(* IEC 61131-3 sources: axsharp/src/ix.blazor/tests/sandbox/ax-blazor-example/src, 40 files *)

(* ---- enumStationStatus.st ---- *)
TYPE enumStationStatus :
    (
        Unknown,
        Available,
        UnAvailable
    );
    END_TYPE

(* ---- stTestEnum.st ---- *)
TYPE stTestEnum :
    (
        Unknown,
        Available,
        UnAvailable
    );
END_TYPE

(* ---- CU00x.st ---- *)
CLASS CU00x EXTENDS CUBase
    VAR PUBLIC
        _cuName: STRING;
    END_VAR
END_CLASS

CLASS CUBase
    VAR PUBLIC
        _baseName : STRING;
    END_VAR
END_CLASS

(* ---- fbWorldWeatherWatch.st ---- *)
CLASS fbWorldWeatherWatch
    VAR PUBLIC
        {#ix-attr:[Container(Layout.Stack)]}
        {#ix-set:AttributeName = "North pole station"}
        //{#ix-set:OpenMap = "https://www.openstreetmap.org/?mlat=74.652&mlon=-95.556#map=6/74.652/-95.556"}
        NorthPole : structWeatherStation := (StationICAO := 'CYRB');
        {#ix-attr:[Container(Layout.Stack)]}
        {#ix-set:AttributeName = "South pole station"}
        //{#ix-set:OpenMap = "https://www.openstreetmap.org/?mlat=-85.05113&mlon=-16.80701#map=1/-85.05113/-16.80701"}
        SouthPole : structWeatherStation := (StationICAO := 'NZSP');
        {#ix-attr:[Container(Layout.Stack)]}
        {#ix-set:AttributeName = "Verl, Germany"}
        //{#ix-set:OpenMap = "https://www.openstreetmap.org/?mlat=51.5799&mlon=8.415#map=6/51.5799/8.4155"}
        Verl : structWeatherStation := (StationICAO := 'EDLP');
        {#ix-attr:[Container(Layout.Stack)]}
        {#ix-set:AttributeName = "Kriva, Slovakia"}
        //{#ix-set:OpenMap = "https://www.openstreetmap.org/?mlat=48.1723&mlon=17.2158#map=6/48.1723/17.2158"}
        Kriva : structWeatherStation := (StationICAO := 'LZIB');
    END_VAR

END_CLASS

(* ---- GroupBox_other.st ---- *)
CLASS GroupBox_other
    VAR PUBLIC
        {#ix-set:AttributeName = "B1"}
        B1: INT;

        {#ix-attr:[Container(Layout.Stack)]}
        {#ix-set:AttributeName = "B2"}
        B2: INT;

        {#ix-attr:[Container(Layout.Stack)]}
        {#ix-set:AttributeName = "A1"}
        Piston_A1 : STRING;
        {#ix-set:AttributeName = "A2"}
        Piston_A2 : STRING;
        {#ix-set:AttributeName = "A3"}
        Piston_A3 : STRING;
        {#ix-set:AttributeName = "A4"}
        Piston_A4 : STRING;

        {#ix-attr:[Container(Layout.Tabs)]}
        Piston_A21 : INT;
        {#ix-set:AttributeName = "A5"}
        Piston_A22 : INT;
        {#ix-set:AttributeName = "A6"}
        Piston_A23 : INT;
        {#ix-set:AttributeName = "A7"}
        Piston_A24 : INT;

        {#ix-attr:[Container(Layout.UniformGrid)]}
        Piston_A31 : REAL;
        {#ix-set:AttributeName = "A8"}
        Piston_A32 : REAL;
        {#ix-set:AttributeName = "A9"}
        Piston_A33 : REAL;
        {#ix-set:AttributeName = "A10"}
        Piston_A34 : REAL;

        Piston_A41 : BOOL;
        {#ix-set:AttributeName = "A11"}
        Piston_A42 : BOOL;
        {#ix-set:AttributeName = "A12"}
        Piston_A43 : BOOL;
        {#ix-set:AttributeName = "A13"}
        Piston_A44 : BOOL;
        {#ix-set:AttributeName = "Servo S1"}
        Servo_S1: TestStructOneGroupWithLayout;
        {#ix-attr:[Container(Layout.Stack)]}
        {#ix-set:AttributeName = "ABB S2"}
        Servo_S2: STRING;
    END_VAR

END_CLASS

(* ---- MAIN.st ---- *)
CLASS MAIN
    VAR PUBLIC
        {#ix-set:AttributeName = "<#Hello#> <#World#>"}
        Hello_World : STRING := 'Hello world!';
        {#ix-set:AttributeName = "cislo"}
        cislo : INT;
        {#ix-set:AttributeName = "bool_val"}
        boolValue : BOOL;
        {#ix-set:AttributeName = "Position"}
        Position : LREAL;
        {#ix-set:AttributeName = "Struct"}
        instanceOfstTest: stTest;
        {#ix-set:AttributeName = "Struct2"}
        instanceOfstTest2: stTest2 ;
        {#ix-set:AttributeName = "instanceOfStTest3"}
        instanceOfstTest3: stTest3 ;
        {#ix-set:AttributeName = "BlazorStruct"}
        instanceOfstBlazor: stBlazor := (testInteger := 10, testString := 'ahoj');
        arr1 : ARRAY [0..2] OF stTest := [(p1 := 6, p2 := 3),(p1 := 9, p2 := 10),(p1 := 12,p2 := 33)];
        arr2 :ARRAY [0..5] OF INT;
        dateVar : DATE;

        {#ix-set:AttributeName = "instanceOfComplex"}
        instanceOfstComplex: stComplex ;
        {#ix-set:AttributeName = "instanceOfStPrimitive"}
        instanceOfstPrimitive: stTestPrimitive ;

    //	{#ix [Container(Layout.Stack)]}
        instanceOfstMultipleLayouts: stMultipleLayouts ;
        instanceOfstMultipleLayouts2: stLayouts ;

        {#ix-set:AttributeName = "instanceOfIxComponent"}
        instanceOfIxComponent: IxComponent ;

        groupBox_test: GroupBox_other;
        cu00: CU00x;
        cuBase: CUBase;
    END_VAR

END_CLASS

(* ---- prgWeatherStations.st ---- *)
{#ix-attr:[Container(Layout.Stack)]}
CLASS prgWeatherStations
    VAR PUBLIC
        {#ix-attr:[Container(Layout.Tabs)]}
        {#ix-set:AttributeName = "Weather Cyclic"}
        _weatherStations : fbWorldWeatherWatch;
        {#ix-attr:[Container(Layout.Stack)]}
        {#ix-attr:[Group(GroupLayout.GroupBox)]}
        {#ix-set:AttributeName = "What plc says"}
        PlcCommentOnCurrentWeather : STRING[254] := 'TEST';
    END_VAR
END_CLASS

(* ---- stBlazor.st ---- *)
CLASS stBlazor
    VAR PUBLIC
        {#ix-set:AttributeName = "<#Integer From PLC#>"}
        testInteger : INT;
        {#ix-set:AttributeName = "testEnum"}
        testEnum : stTestEnum;
        {#ix-set:AttributeName = "<#String From PLC#>"}
        testString : STRING;
        testReal : REAL := REAL#592.25;
        {#ix-attr:[RenderIgnore("Display")]}
        testLReal : LREAL := 42.2;
        testBool : BOOL;
        {#ix-set:AttributeName = "Complex"}
        {#ix-attr:[RenderIgnore()]}
        complexInstance : stComplex := (stComplexInteger := 33, stComplexString := 'hello world');
        {#ix-set:AttributeName = "testInstance1"}
        testInstance : stTest3;
        {#ix-set:AttributeName = "testInstance2"}
        testInstance2 : stTest3;
        {#ix-set:AttributeName = "testInstance3"}
        testInstance3 : stTest;
    END_VAR

END_CLASS

(* ---- stComplex.st ---- *)
CLASS stComplex
    VAR PUBLIC
        {#ix-set:AttributeName = "<#Integer From PLC#>"}
        stComplexInteger : INT;
        {#ix-set:AttributeName = "<#String From PLC#>"}
        stComplexString : STRING;
    END_VAR

END_CLASS

(* ---- stComplexUnknown.st ---- *)
CLASS stComplexUnknown
    VAR PUBLIC
        {#ix-set:AttributeName = "<#String unknown From PLC#>"}
        stComplexUnknownString : STRING;
        {#ix-set:AttributeName = "<#BOOL unknown From PLC#>"}
        testBool : BOOL;
        {#ix-set:AttributeName = "<#Integer unknown From PLC#>"}
        stComplexUnknowInteger : INT;
        {#ix-set:AttributeName = "<#DATE unknown From PLC#>"}
        TestDate : DATE;
    END_VAR
END_CLASS

(* ---- stExample.st ---- *)
CLASS stExample
    VAR PUBLIC
        {#ix-attr:[Container(Layout.Tabs)]}
        {#ix-attr:[Group(GroupLayout.GroupBox)]}
        {#ix-set:AttributeName = "Group name"}
        testInteger : INT;
        testEnum : stTestEnum;
        testString : STRING := 'Hello World';
        testBool : BOOL;
    END_VAR

END_CLASS

(* ---- stLayouts.st ---- *)
CLASS stLayouts
    VAR
        {#ix-set:AttributeName = "B1"}
	B1: INT;

	{#ix-attr:[Container(Layout.Stack)]}
	{#ix-set:AttributeName = "B2"}
	B2: INT;

	{#ix-attr:[Container(Layout.Stack)]}
	{#ix-set:AttributeName = "A1"}
	Piston_A1 : STRING;
	{#ix-set:AttributeName = "A2"}
	Piston_A2 : STRING;
	{#ix-set:AttributeName = "A3"}
	Piston_A3 : STRING;
	{#ix-set:AttributeName = "A4"}
	Piston_A4 : STRING;

	{#ix-attr:[Container(Layout.Tabs)]}
	Piston_A21 : INT;
	{#ix-set:AttributeName = "A5"}
	Piston_A22 : INT;
	{#ix-set:AttributeName = "A6"}
	Piston_A23 : INT;
	{#ix-set:AttributeName = "A7"}
	Piston_A24 : INT;

	{#ix-attr:[Container(Layout.UniformGrid)]}
	Piston_A31 : REAL;
	{#ix-set:AttributeName = "A8"}
	Piston_A32 : REAL;
	{#ix-set:AttributeName = "A9"}
	Piston_A33 : REAL;
	{#ix-set:AttributeName = "A10"}
	Piston_A34 : REAL;

	Piston_A41 : BOOL;
	{#ix-set:AttributeName = "A11"}
	Piston_A42 : BOOL;
	{#ix-set:AttributeName = "A12"}
	Piston_A43 : BOOL;
	{#ix-set:AttributeName = "A13"}
	Piston_A44 : BOOL;

	{#ix-set:AttributeName = "Servo S1"}
	Servo_S1: TestStructOneGroupWithLayout;
	{#ix-attr:[Container(Layout.Stack)]}
	{#ix-set:AttributeName = "ABB S2"}
	Servo_S2: STRING;
    END_VAR
END_CLASS

(* ---- stMultipleLayouts.st ---- *)
CLASS stMultipleLayouts
    VAR PUBLIC
        {#ix-attr:[Container(Layout.Tabs)]}
        {#ix-set:AttributeName = "With One Group Layout"}
        Servo_S5: TestStructOneGroupWithLayout;

        {#ix-attr:[Container(Layout.Tabs)]}
        {#ix-set:AttributeName = "Without Group Layout"}
        Servo_S6: TestStruct;

        {#ix-attr:[Container(Layout.Tabs)]}
        {#ix-set:AttributeName = "With Multiple Groups "}
        Servo_S7: TestStructMultipleGroups;

        {#ix-attr:[Container(Layout.Tabs)]}
        {#ix-set:AttributeName = "TestStruct With Main Layout  "}
        Servo_S8: TestStructWithMainLayout;

        {#ix-attr:[Container(Layout.Stack)]}
        {#ix-set:AttributeName = "A1"}
        Piston_A1 : STRING;
        {#ix-set:AttributeName = "A2"}
        Piston_A2 : STRING;
        {#ix-set:AttributeName = "A3"}
        Piston_A3 : STRING;
        {#ix-set:AttributeName = "A4"}
        Piston_A4 : STRING;

        {#ix-attr:[Container(Layout.Wrap)]}
        {#ix-set:AttributeName = "A5"}
        Piston_A21 : INT;
        {#ix-set:AttributeName = "A6"}
        Piston_A22 : INT;
        {#ix-set:AttributeName = "A7"}
        Piston_A23 : INT;
        {#ix-set:AttributeName = "A8"}
        Piston_A24 : INT;

        {#ix-attr:[Container(Layout.Tabs)]}
        Piston_A31 : REAL;
        {#ix-set:AttributeName = "A8"}
        Piston_A32 : REAL;
        {#ix-set:AttributeName = "A9"}
        Piston_A33 : REAL;
        {#ix-set:AttributeName = "A10"}
        Piston_A34 : REAL;

        {#ix-attr:[Container(Layout.UniformGrid)]}
        Piston_A41 : BOOL;
        {#ix-set:AttributeName = "A11"}
        Piston_A42 : BOOL;
        {#ix-set:AttributeName = "A12"}
        Piston_A43 : BOOL;
        {#ix-set:AttributeName = "A13"}
        Piston_A44 : BOOL;

        {#ix-attr:[Container(Layout.Stack)]}
        {#ix-set:AttributeName = "Servo S1"}
        Servo_S1: STRING;

        {#ix-attr:[Container(Layout.Stack)]}
        {#ix-set:AttributeName = "ABB S2"}
        Servo_S2: STRING;

        {#ix-attr:[Container(Layout.Tabs)]}
        {#ix-set:AttributeName = "My ix component"}
        component: IxComponent;
        {#ix-set:AttributeName = "Servo S3"}
        Servo_S3: stTest3;
        {#ix-set:AttributeName = "Servo S4"}
        Servo_S4: stTest3;

    END_VAR

END_CLASS

(* ---- structWeatherStation.st ---- *)
CLASS structWeatherStation
    VAR PUBLIC
        {#ix-set:AttributeName = "Station name (ICAO)"}
        StationICAO : STRING[4];
        {#ix-set:AttributeName = "Station status"}
        StationStatus : enumStationStatus;
        {#ix-set:AttributeName = "Dew Point"}
        {#ix-set:AttributeUnits = "°C"}
        {#ix-attr:[RenderIgnore()]}
        DewPoint : REAL;
        {#ix-set:AttributeName = "Pressure"}
        {#ix-set:AttributeUnits = "Torr"}
        Pressure : REAL;
        {#ix-set:AttributeName = "Temperature"}
        {#ix-set:AttributeUnits = "°C"}
        Temp : REAL;
        {#ix-set:AttributeName = "Visibility"}
        {#ix-set:AttributeUnits = "km"}
        Visibility : REAL;
        {#ix-set:AttributeName = "Wind heading"}
        {#ix-set:AttributeUnits = "Azimuth"}
        WindHeading : UINT;
        {#ix-set:AttributeName = "Wind speed"}
        {#ix-set:AttributeUnits = "m/s"}
        WindSpeed : REAL;
        TestDate : DATE;
        TestDateTime : DATE_AND_TIME;
        TestTimeOfDay : TIME_OF_DAY;
    END_VAR

END_CLASS

(* ---- stSimplePrimitive.st ---- *)
CLASS stSimplePrimitive
    VAR PUBLIC
        {#ix-set:AttributeName = "<#Test Integer#>"}
        testInteger : INT;
        {#ix-set:AttributeName = "<#Test String#>"}
        testString : STRING;
    END_VAR
END_CLASS

(* ---- stTest.st ---- *)
CLASS stTest
    VAR PUBLIC
        p1:INT;
        p2:INT;
        stTest3Struct: stTest3;
        DateVar2: DATE;
        complexInstanceNested : stComplex := (stComplexInteger := 13, stComplexString := 'hello nested');
    END_VAR

END_CLASS

(* ---- stTest2.st ---- *)
CLASS stTest2
    VAR
        testVarString: STRING;
        testVarInt: INT;
        instanceOfstTest3: stTest3;
        arr1 : ARRAY [0..2] OF stTest := [(p1 := 445, p2 := 446),(p1 := 152, p2 := 100),(p1 := 121,p2 := 338)];
    END_VAR

END_CLASS

(* ---- stTest3.st ---- *)
CLASS stTest3
    VAR PUBLIC
        ix_bool : BOOL;
        ix_int : INT;
        ix_string : STRING;
    END_VAR
END_CLASS

(* ---- stTestComplex.st ---- *)
CLASS stTestComplex
    VAR PUBLIC
        {#ix-set:AttributeName = "<#Integer From PLC#>"}
        testInteger : INT;
        {#ix-set:AttributeName = "<#Complex Instance#>"}
        testComplexInstance : stComplex := (stComplexInteger := 33, stComplexString := 'hello world');
        {#ix-set:AttributeName = "<#String From PLC#>"}
        testString : STRING;
        {#ix-attr:[Container(Layout.Stack)]}
        {#ix-set:AttributeName = "<#Complex Instance#>"}
        testComplexUnknownInstance : stComplexUnknown;
    END_VAR

END_CLASS

(* ---- stTestLayouts.st ---- *)
CLASS stTestLayouts
    VAR PUBLIC
        {#ix-attr:[Container(Layout.Stack)]}
        test_stack: stSimplePrimitive;
        {#ix-attr:[Container(Layout.Wrap)]}
        test_wrap: stSimplePrimitive;
        {#ix-attr:[Container(Layout.Tabs)]}
        test_tabs: stSimplePrimitive;
        {#ix-attr:[Container(Layout.UniformGrid)]}
        test_uniform: stSimplePrimitive;

        {#ix-attr:[Container(Layout.Stack)]}
        {#ix-attr:[Group(GroupLayout.GroupBox)]}
        test_groupbox_stack: stSimplePrimitive;

        {#ix-attr:[Container(Layout.Stack)]}
        {#ix-attr:[Group(GroupLayout.Border)]}
        test_border_stack: stSimplePrimitive;

        {#ix-attr:[Container(Layout.Wrap)]}
        {#ix-attr:[Group(GroupLayout.GroupBox)]}
        test_groupbox_wrap: stSimplePrimitive;

        {#ix-attr:[Container(Layout.Wrap)]}
        {#ix-attr:[Group(GroupLayout.Border)]}
        test_border_wrap: stSimplePrimitive;

        {#ix-attr:[Container(Layout.Tabs)]}
        {#ix-attr:[Group(GroupLayout.GroupBox)]}
        test_groupbox_tabs: stSimplePrimitive;

        {#ix-attr:[Container(Layout.Tabs)]}
        {#ix-attr:[Group(GroupLayout.Border)]}
        test_border_tabs: stSimplePrimitive;

        {#ix-attr:[Container(Layout.UniformGrid)]}
        {#ix-attr:[Group(GroupLayout.GroupBox)]}
        test_groupbox_uniformGrid: stSimplePrimitive;

        {#ix-attr:[Container(Layout.UniformGrid)]}
        {#ix-attr:[Group(GroupLayout.Border)]}
        test_border_uniformGrid: stSimplePrimitive;
    END_VAR
END_CLASS

(* ---- stTestMultipleNested.st ---- *)
CLASS stTestMultipleNested
    VAR PUBLIC
        {#ix-attr:[Container(Layout.Tabs)]}
        {#ix-set:AttributeName = "With One Group Layout"}
        Servo_S5: TestStructOneGroupWithLayout;

        {#ix-attr:[Container(Layout.Tabs)]}
        {#ix-set:AttributeName = "Without Group Layout"}
        Servo_S6: TestStruct;

        {#ix-attr:[Container(Layout.Tabs)]}
        {#ix-set:AttributeName = "With Multiple Groups "}
        Servo_S7: TestStructMultipleGroups;

        {#ix-attr:[Container(Layout.Tabs)]}
        {#ix-set:AttributeName = "TestStruct With Main Layout  "}
        Servo_S8: TestStructWithMainLayout;

        {#ix-attr:[Container(Layout.Stack)]}
        {#ix-set:AttributeName = "A1"}
        Piston_A1 : STRING;
        {#ix-set:AttributeName = "A2"}
        Piston_A2 : STRING;
        {#ix-set:AttributeName = "A3"}
        Piston_A3 : STRING;
        {#ix-set:AttributeName = "A4"}
        Piston_A4 : STRING;

        {#ix-attr:[Container(Layout.Wrap)]}
        {#ix-set:AttributeName = "A5"}
        Piston_A21 : INT;
        {#ix-set:AttributeName = "A6"}
        Piston_A22 : INT;
        {#ix-set:AttributeName = "A7"}
        Piston_A23 : INT;
        {#ix-set:AttributeName = "A8"}
        Piston_A24 : INT;

        {#ix-attr:[Container(Layout.Tabs)]}
        Piston_A31 : REAL;
        {#ix-set:AttributeName = "A8"}
        Piston_A32 : REAL;
        {#ix-set:AttributeName = "A9"}
        Piston_A33 : REAL;
        {#ix-set:AttributeName = "A10"}
        Piston_A34 : REAL;

        {#ix-attr:[Container(Layout.UniformGrid)]}
        Piston_A41 : BOOL;
        {#ix-set:AttributeName = "A11"}
        Piston_A42 : BOOL;
        {#ix-set:AttributeName = "A12"}
        Piston_A43 : BOOL;
        {#ix-set:AttributeName = "A13"}
        Piston_A44 : BOOL;

        {#ix-attr:[Container(Layout.Stack)]}
        {#ix-set:AttributeName = "Servo S1"}
        Servo_S1: STRING;

        {#ix-attr:[Container(Layout.Stack)]}
        {#ix-set:AttributeName = "ABB S2"}
        Servo_S2: STRING;

        {#ix-attr:[Container(Layout.Tabs)]}
        {#ix-set:AttributeName = "My ix component"}
        component: IxComponent;
        {#ix-set:AttributeName = "Servo S3"}
        Servo_S3: STRING;
        {#ix-set:AttributeName = "Servo S4"}
        Servo_S4: STRING;
    END_VAR

END_CLASS

(* ---- stTestNested.st ---- *)
CLASS stTestNested
    VAR PUBLIC
        {#ix-attr:[Container(Layout.Wrap)]}
        e:INT;
        r44:STRING;
        k21:STRING;
    END_VAR

END_CLASS

(* ---- stTestPrimitive.st ---- *)
CLASS stTestPrimitive
    VAR PUBLIC
        {#ix-set:AttributeName = "<#Integer From PLC#>"}
        testInteger : INT;
        {#ix-set:AttributeName = "<#UInteger From PLC#>"}
        testUInteger : INT;
        {#ix-set:AttributeName = "<#STRING From PLC#>"}
        testString : STRING;
        {#ix-set:AttributeName = "<#WORD From PLC#>"}
        testWord : WORD;
        {#ix-set:AttributeName = "<#BYTE From PLC#>"}
        testByte : BYTE;
        {#ix-set:AttributeName = "<#REAL From PLC#>"}
        testReal : REAL;
        {#ix-set:AttributeName = "<#LREAL From PLC#>"}
        testLReal : LREAL;
        {#ix-set:AttributeName = "<#BOOL From PLC#>"}
        testBool : BOOL;
        {#ix-set:AttributeName = "<#DATE From PLC#>"}
        TestDate : DATE;
        {#ix-set:AttributeName = "<#DATE_AND_TIME From PLC#>"}
        TestDateTime : DATE_AND_TIME;
        {#ix-set:AttributeName = "<#TIME_OF_DAY From PLC#>"}
        TestTimeOfDay : TIME_OF_DAY;
    END_VAR

END_CLASS

(* ---- stTestRenderIgnore.st ---- *)
CLASS stTestRenderIgnore
    VAR PUBLIC
        {#ix-attr:[RenderIgnore()]}
        {#ix-set:AttributeName = "<#Integer From PLC#>"}
        testInteger : INT;
        {#ix-set:AttributeName = "<#UInteger From PLC#>"}
        testUInteger : INT;
        {#ix-set:AttributeName = "<#STRING From PLC#>"}
        testString : STRING;
        {#ix-set:AttributeName = "<#WORD From PLC#>"}
        testWord : WORD;
        {#ix-set:AttributeName = "<#BYTE From PLC#>"}
        testByte : BYTE;
        {#ix-set:AttributeName = "<#REAL From PLC#>"}
        testReal : REAL;
        {#ix-set:AttributeName = "<#LREAL From PLC#>"}
        testLReal : LREAL;
        {#ix-attr:[RenderIgnore("Display","ShadowDisplay")]}
        {#ix-set:AttributeName = "<#BOOL From PLC#>"}
        testBool : BOOL;
        {#ix-attr:[RenderIgnore("Control","ShadowControl")]}
        {#ix-set:AttributeName = "<#DATE From PLC#>"}
        TestDate : DATE;
        {#ix-set:AttributeName = "<#DATE_AND_TIME From PLC#>"}
        TestDateTime : DATE_AND_TIME;
    END_VAR

END_CLASS

(* ---- TcoVortexObject.st ---- *)
CLASS TcoIxObject
    VAR PUBLIC
        ix_bool : BOOL;
        ix_int : INT;
        ix_string : STRING;
    END_VAR
END_CLASS

(* ---- TestEmpty.st ---- *)
CLASS TestEmpty
    VAR PUBLIC

    END_VAR

END_CLASS

(* ---- testingProgram.st ---- *)
CLASS testingProgram
    VAR PUBLIC
        {#ix-set:AttributeName = "instanceOfStPrimitive"}
        {#ix-attr:[Container(Layout.Wrap)]}
        testPrimitive: stTestPrimitive;
        {#ix-set:AttributeName = "instanceOfStPrimitive"}
        testComplex: stTestComplex;
        {#ix-set:AttributeName = "instanceOfStEnum"}
        testEnum: stTestEnum;
        {#ix-attr:[Container(Layout.UniformGrid)]}
        testRenderIgnore : stTestRenderIgnore;

        testEmpty: TestEmpty;
        testLayoutOverwrite: TestLayoutOverwriting;
        testMixed : TestMixed;
        testMultipleLayouts: TestMultipleLayouts;
        testSimple: TestSimple;
        testWithoutLayouts: TestWithoutLayouts;
        testSimpleNested: TestSimpleNested;
        {#ix-attr:[Container(Layout.Tabs)]}
        testMultipleNested: stTestMultipleNested;

        testLayouts : stTestLayouts;
    END_VAR

END_CLASS

(* ---- TestLayoutOverwriting.st ---- *)
{#ix-attr:[Container(Layout.UniformGrid)]}
CLASS TestLayoutOverwriting
    VAR PUBLIC
        ix_bool : BOOL;
        ix_int : INT;
        ix_string : STRING;

        {#ix-attr:[Container(Layout.Wrap)]}
        simple: TestSimple;

        {#ix-attr:[Container(Layout.Wrap)]}
        weather: prgWeatherStations;
    END_VAR

END_CLASS

(* ---- TestMixed.st ---- *)
CLASS TestMixed
    VAR PUBLIC
        {#ix-attr:[Container(Layout.Wrap)]}
        e:INT;
        r44:STRING;
        k21:STRING;
    END_VAR
END_CLASS

(* ---- TestMultipleLayouts.st ---- *)
CLASS TestMultipleLayouts
    VAR PUBLIC
        {#ix-set:AttributeName = "B1"}
        B1: INT;

        {#ix-attr:[Container(Layout.Stack)]}
        {#ix-set:AttributeName = "B2"}
        B2: INT;

        {#ix-attr:[Container(Layout.Stack)]}
        {#ix-set:AttributeName = "A1"}
        Piston_A1 : STRING;
        {#ix-set:AttributeName = "A2"}
        Piston_A2 : STRING;
        {#ix-set:AttributeName = "A3"}
        Piston_A3 : STRING;
        {#ix-set:AttributeName = "A4"}
        Piston_A4 : STRING;

        {#ix-attr:[Container(Layout.Tabs)]}
        Piston_A21 : INT;
        {#ix-set:AttributeName = "A5"}
        Piston_A22 : INT;
        {#ix-set:AttributeName = "A6"}
        Piston_A23 : INT;
        {#ix-set:AttributeName = "A7"}
        Piston_A24 : INT;

        {#ix-attr:[Container(Layout.UniformGrid)]}
        Piston_A31 : REAL;
        {#ix-set:AttributeName = "A8"}
        Piston_A32 : REAL;
        {#ix-set:AttributeName = "A9"}
        Piston_A33 : REAL;
        {#ix-set:AttributeName = "A10"}
        Piston_A34 : REAL;

        Piston_A41 : BOOL;
        {#ix-set:AttributeName = "A11"}
        Piston_A42 : BOOL;
        {#ix-set:AttributeName = "A12"}
        Piston_A43 : BOOL;
        {#ix-set:AttributeName = "A13"}
        Piston_A44 : BOOL;
        {#ix-attr:[Container(Layout.Stack)]}
        {#ix-set:AttributeName = "Servo S1"}
        Servo_S1: STRING;
        {#ix-attr:[Container(Layout.Stack)]}
        {#ix-set:AttributeName = "ABB S2"}
        Servo_S2: STRING;
    END_VAR

END_CLASS

(* ---- TestSimple.st ---- *)
CLASS TestSimple
    VAR PUBLIC
        {#ix-set:AttributeName = "A1"}
        Piston_A1 : STRING;
        {#ix-set:AttributeName = "A2"}
        Piston_A2 : STRING;
        {#ix-set:AttributeName = "A3"}
        Piston_A3 : STRING;
        {#ix-set:AttributeName = "A4"}
        Piston_A4 : STRING;
    END_VAR
END_CLASS

(* ---- TestSimpleNested.st ---- *)
CLASS TestSimpleNested
    VAR PUBLIC
        {#ix-attr:[Container(Layout.Tabs)]}
	    str: stTestNested;
    END_VAR

END_CLASS

(* ---- TestStruct.st ---- *)
CLASS TestStruct
    VAR PUBLIC
        e:INT;
        r44:STRING;
        k21:STRING;
        example:stExample;
    END_VAR

END_CLASS

(* ---- TestStructMultipleGroups.st ---- *)
CLASS TestStructMultipleGroups
    VAR PUBLIC
        e:INT;
        {#ix-attr:[Container(Layout.Stack)]}
        r44:STRING;
        k21:STRING;
    END_VAR

END_CLASS

(* ---- TestStructOneGroupWithLayout.st ---- *)
CLASS TestStructOneGroupWithLayout
    VAR PUBLIC
        {#ix-attr:[Container(Layout.Wrap)]}
        e:INT;
        r44:STRING;
        k21:STRING;
    END_VAR

END_CLASS

(* ---- TestStructWithMainLayout.st ---- *)
CLASS TestStructWithMainLayout
    VAR PUBLIC
        e:INT;
        r44:STRING;
        k21:STRING;
    END_VAR
END_CLASS

(* ---- TestWithoutLayouts.st ---- *)
CLASS TestWithoutLayouts
    VAR PUBLIC
        ix_bool : BOOL;
        ix_int : INT;
        ix_string : STRING;
    END_VAR

END_CLASS

(* ---- VortexComponents.st ---- *)
CLASS IxComponent
    VAR PUBLIC
        ix_bool : BOOL;
        ix_int : INT;
        ix_string : STRING;
    END_VAR
END_CLASS

(* ---- configuration.st ---- *)
CONFIGURATION MyConfiguration
    TASK Main(Interval := T#1000ms, Priority := 1);
    PROGRAM P1 WITH Main: MyProgram;

    VAR_GLOBAL
        testingProgram : testingProgram;
        prgWeatherStations : prgWeatherStations;
        MAINC : MAIN;
    END_VAR
END_CONFIGURATION

(* ---- program.st ---- *)
PROGRAM MyProgram
    VAR_EXTERNAL

    END_VAR

    VAR

    END_VAR

    VAR_TEMP

    END_VAR

    // code here
    ;
END_PROGRAM
